// TIA Portal V20 export
// export: Created 2026-10-31T19:03:51.7054379Z, ExportSetting WithDefaults, WithReadOnly
Screen "zzTestControls"  1280x800, Number=3
  ScreenLayer 
    UserView "User view_1" at 13,309 size 480x240  Appearance=AppearanceFlat, CountVisibleItems=8, ViewType=ViewTypeComplex
